FUNCTION_BLOCK FB_Unit
VAR_INPUT
END_VAR
VAR_OUTPUT
END_VAR
VAR
END_VAR

END_FUNCTION_BLOCK

(* stored: Version 1.1.0.1
   POU FB_Unit: Id {0ac84c1d-b47a-41f1-a8f9-f65828d55eaa}, SpecialFunc None *)
